SUBAPPLICATION OptionalGroup_002a (* Optionsgruppe 2a: wie OptionalGroup_001a, aber mit Input_I2/Output_Q2 - Gegenstueck mit Plug AOption_OUT zu OptionalGroup_002; wie OptionalGroup_001b (Eingang/Ausgang per QI freigeschaltet), reicht die Aktivierung zusaetzlich ueber den Plug AOption_OUT an eine nachgeschaltete Gruppe weiter - fuer sequenzielle Aktivierung mehrerer Gruppen (erst 2a, dann nachgeschaltete Gruppe). *)
  (* Standard: 61499-2; Description: Copyright (c) 2026 Meisterschulen am Ostbahnhof This program and the accompanying materials are made available under the terms of the Eclipse Public License 2.0 which is available at https://www.eclipse.org/legal/epl-2.0/ SPDX-License-Identifier: EPL-2.0 *)
  (* Version 1.0, 2026-10-17, Franz Höpfinger, Meisterschulen am Ostbahnhof, Baugleich zu OptionalGroup_001a mit I2/Q2. Daisy-Chain-Glied fuer sequenzielle Options-Aktivierung: AOption_OUT (Option::AOption) wird erst ausgeloest, wenn DigitalOutput_Q2 selbst initialisiert ist, und dessen INIT_CNF wird an den eigenen Socket AOption_IN zurueckgemeldet - der aufrufende DEMUX sieht die Gruppe also erst als fertig, wenn die GESAMTE Kette (inkl. nachgeschalteter Gruppen an AOption_OUT) bestaetigt hat. *)
  PACKAGE MyLib_AX_Option::sys;
  IMPORT logiBUS::io::DI::logiBUS_DI::Input_I2;
  IMPORT logiBUS::io::DQ::logiBUS_DO::Output_Q2;
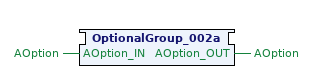
  SOCKETS
    AOption_IN : Option::AOption;
  END_SOCKETS
  PLUGS
    AOption_OUT : Option::AOption;
  END_PLUGS
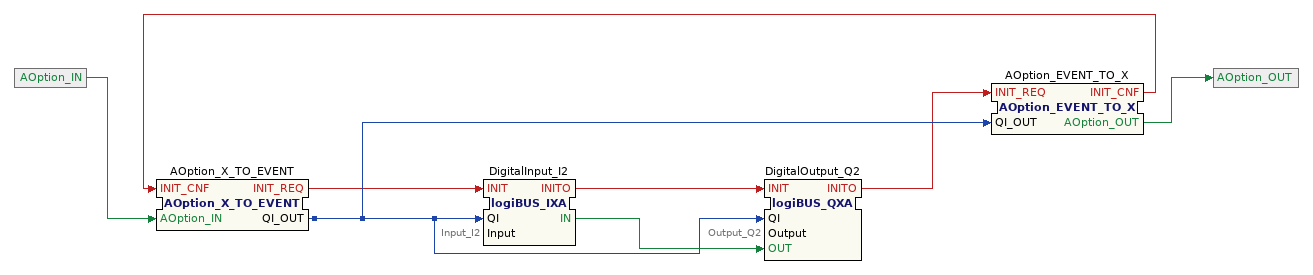
  FBS
    DigitalInput_I2 : logiBUS::io::DI::logiBUS_IXA(Input := Input_I2);
    DigitalOutput_Q2 : logiBUS::io::DQ::logiBUS_QXA(Output := Output_Q2);
    AOption_X_TO_EVENT : Option::conversion::AOption_X_TO_EVENT;
    AOption_EVENT_TO_X : Option::conversion::AOption_EVENT_TO_X;
  END_FBS
  EVENT_CONNECTIONS
    AOption_X_TO_EVENT.INIT_REQ TO DigitalInput_I2.INIT;
    DigitalInput_I2.INITO TO DigitalOutput_Q2.INIT;
    DigitalOutput_Q2.INITO TO AOption_EVENT_TO_X.INIT_REQ;
    AOption_EVENT_TO_X.INIT_CNF TO AOption_X_TO_EVENT.INIT_CNF;
  END_CONNECTIONS
  DATA_CONNECTIONS
    AOption_X_TO_EVENT.QI_OUT TO DigitalInput_I2.QI;
    AOption_X_TO_EVENT.QI_OUT TO DigitalOutput_Q2.QI;
    AOption_X_TO_EVENT.QI_OUT TO AOption_EVENT_TO_X.QI_OUT;
  END_CONNECTIONS
  ADAPTER_CONNECTIONS
    DigitalInput_I2.IN TO DigitalOutput_Q2.OUT;
    AOption_IN TO AOption_X_TO_EVENT.AOption_IN;
    AOption_EVENT_TO_X.AOption_OUT TO AOption_OUT;
  END_CONNECTIONS
END_SUBAPPLICATION
